FUNCTION_BLOCK Sensor_Generico_HMI (* Service Interface Function Block Type *)
  (* Standard: 61499-2 *)
  (* Version 1.6, 12/11/2026, Hidryco, Hidryco, 1.6: STS_CODIGO_ERRO, STS_CODIGO_AVISO e STS_ALM_AVISO_EST (aviso/erro do proprio dispositivo). 1.5: CommonError, Reliability e DaysToMaintenance para a IO List da Nereda. 1.4: STS_LIMITE_HH..LL (limites dos alarmes em unidade de engenharia) para o grafico. IHM do Sensor_Generico *)
  PACKAGE Hidryco.HidrycoLib;
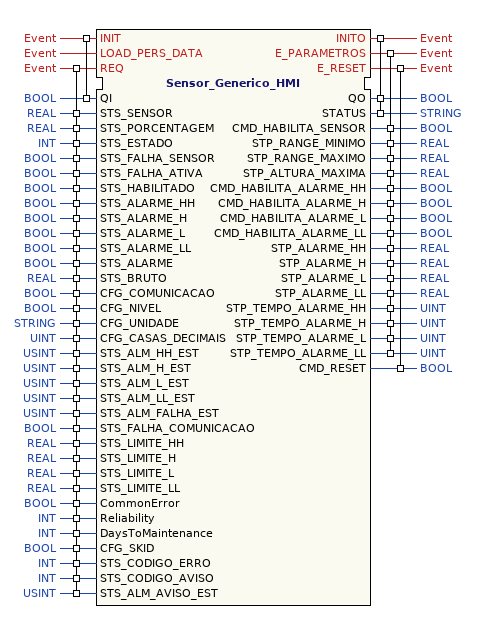
  EVENT_INPUT
    INIT WITH QI;
    LOAD_PERS_DATA; (* Reenvia os parametros persistentes *)
    REQ WITH STS_SENSOR, STS_PORCENTAGEM, STS_ESTADO, STS_FALHA_SENSOR, STS_FALHA_ATIVA, STS_HABILITADO, STS_ALARME_HH, STS_ALARME_H, STS_ALARME_L, STS_ALARME_LL, STS_ALARME, STS_BRUTO, CFG_COMUNICACAO, CFG_NIVEL, CFG_UNIDADE, CFG_CASAS_DECIMAIS, STS_ALM_HH_EST, STS_ALM_H_EST, STS_ALM_L_EST, STS_ALM_LL_EST, STS_ALM_FALHA_EST, STS_FALHA_COMUNICACAO, STS_LIMITE_HH, STS_LIMITE_H, STS_LIMITE_L, STS_LIMITE_LL, CommonError, Reliability, DaysToMaintenance, CFG_SKID, STS_CODIGO_ERRO, STS_CODIGO_AVISO, STS_ALM_AVISO_EST; (* Atualizacao de status *)
  END_EVENT
  EVENT_OUTPUT
    INITO WITH QO, STATUS;
    E_PARAMETROS WITH CMD_HABILITA_SENSOR, STP_RANGE_MINIMO, STP_RANGE_MAXIMO, STP_ALTURA_MAXIMA, CMD_HABILITA_ALARME_HH, CMD_HABILITA_ALARME_H, CMD_HABILITA_ALARME_L, CMD_HABILITA_ALARME_LL, STP_ALARME_HH, STP_ALARME_H, STP_ALARME_L, STP_ALARME_LL, STP_TEMPO_ALARME_HH, STP_TEMPO_ALARME_H, STP_TEMPO_ALARME_L, STP_TEMPO_ALARME_LL;
    E_RESET WITH CMD_RESET;
  END_EVENT
  VAR_INPUT
    QI : BOOL;
    STS_SENSOR : REAL; (* Valor em unidade de engenharia *) {SET_ATTRIBUTE(Runtime.History.Depth, 500)} {SET_ATTRIBUTE(Runtime.History.SmoothTime, 60000)} {SET_ATTRIBUTE(Runtime.History.SmoothValue, 0.1)}
    STS_PORCENTAGEM : REAL; (* Nivel em % (so sensor de nivel) *)
    STS_ESTADO : INT; (* 0 normal, 1 alerta, 2 alarme, 3 falha, 4 desabilitado *)
    STS_FALHA_SENSOR : BOOL; (* Falha do sensor (4-20 mA fora da faixa ou falha do instrumento), sem a falha de comunicacao *)
    STS_FALHA_ATIVA : BOOL; (* Qualquer falha ativa (sensor ou comunicacao) *)
    STS_HABILITADO : BOOL; (* Sensor habilitado *)
    STS_ALARME_HH : BOOL; (* Alarme HH *)
    STS_ALARME_H : BOOL; (* Alarme H *)
    STS_ALARME_L : BOOL; (* Alarme L *)
    STS_ALARME_LL : BOOL; (* Alarme LL *)
    STS_ALARME : BOOL; (* Algum alarme *)
    STS_BRUTO : REAL; (* Valor bruto lido (diagnostico) *)
    CFG_COMUNICACAO : BOOL; (* Configuracao: valor por comunicacao *)
    CFG_NIVEL : BOOL; (* Configuracao: sensor de nivel (mostra %) *)
    CFG_UNIDADE : STRING; (* Configuracao: unidade de engenharia *)
    CFG_CASAS_DECIMAIS : UINT; (* Configuracao: casas decimais *)
    STS_ALM_HH_EST : USINT; (* Estado do ALARM_BIT HH (0 normal, 1 ativo reconhecido, 2 ativo nao reconhecido, 3 saiu nao reconhecido, 4 ativo e saiu nao reconhecido) *)
    STS_ALM_H_EST : USINT; (* Estado do ALARM_BIT H (0 normal, 1 ativo reconhecido, 2 ativo nao reconhecido, 3 saiu nao reconhecido, 4 ativo e saiu nao reconhecido) *)
    STS_ALM_L_EST : USINT; (* Estado do ALARM_BIT L (0 normal, 1 ativo reconhecido, 2 ativo nao reconhecido, 3 saiu nao reconhecido, 4 ativo e saiu nao reconhecido) *)
    STS_ALM_LL_EST : USINT; (* Estado do ALARM_BIT LL (0 normal, 1 ativo reconhecido, 2 ativo nao reconhecido, 3 saiu nao reconhecido, 4 ativo e saiu nao reconhecido) *)
    STS_ALM_FALHA_EST : USINT; (* Estado do ALARM_BIT FALHA (0 normal, 1 ativo reconhecido, 2 ativo nao reconhecido, 3 saiu nao reconhecido, 4 ativo e saiu nao reconhecido) *)
    STS_FALHA_COMUNICACAO : BOOL; (* Falha de comunicacao do sensor *)
    STS_LIMITE_HH : REAL; (* Limite do alarme HH em unidade de engenharia *) {SET_ATTRIBUTE(Runtime.History.Depth, 100)} {SET_ATTRIBUTE(Runtime.History.SmoothTime, 60000)} {SET_ATTRIBUTE(Runtime.History.SmoothValue, 0)}
    STS_LIMITE_H : REAL; (* Limite do alarme H em unidade de engenharia *) {SET_ATTRIBUTE(Runtime.History.Depth, 100)} {SET_ATTRIBUTE(Runtime.History.SmoothTime, 60000)} {SET_ATTRIBUTE(Runtime.History.SmoothValue, 0)}
    STS_LIMITE_L : REAL; (* Limite do alarme L em unidade de engenharia *) {SET_ATTRIBUTE(Runtime.History.Depth, 100)} {SET_ATTRIBUTE(Runtime.History.SmoothTime, 60000)} {SET_ATTRIBUTE(Runtime.History.SmoothValue, 0)}
    STS_LIMITE_LL : REAL; (* Limite do alarme LL em unidade de engenharia *) {SET_ATTRIBUTE(Runtime.History.Depth, 100)} {SET_ATTRIBUTE(Runtime.History.SmoothTime, 60000)} {SET_ATTRIBUTE(Runtime.History.SmoothValue, 0)}
    CommonError : BOOL; (* Nereda: erro do sensor (= STS_FALHA_SENSOR) *)
    Reliability : INT; (* Nereda: confiabilidade do sensor (%), fixo em 80 *)
    DaysToMaintenance : INT; (* Nereda: dias para a manutencao (sem fonte: 0) *)
    CFG_SKID : BOOL; (* Configuracao: valor ja escalado no skid (sem ajuste de escala na IHM) *)
    STS_CODIGO_ERRO : INT; (* Codigo de erro do proprio dispositivo (0 = nenhum) *)
    STS_CODIGO_AVISO : INT; (* Codigo de aviso do proprio dispositivo (0 = nenhum) *)
    STS_ALM_AVISO_EST : USINT; (* Estado do ALARM_BIT de aviso do dispositivo (0 normal, 1 ativo reconhecido, 2 ativo nao reconhecido, 3 saiu nao reconhecido, 4 ativo e saiu) *)
  END_VAR
  VAR_OUTPUT
    QO : BOOL; (* Event Output Qualifier *)
    STATUS : STRING; (* Service Status *)
    CMD_HABILITA_SENSOR : BOOL; (* Sensor habilitado *)
    STP_RANGE_MINIMO : REAL; (* Valor de engenharia em 4 mA *)
    STP_RANGE_MAXIMO : REAL; (* Valor de engenharia em 20 mA *)
    STP_ALTURA_MAXIMA : REAL; (* Altura maxima do tanque (nivel) *)
    CMD_HABILITA_ALARME_HH : BOOL; (* Alarme HH habilitado *)
    CMD_HABILITA_ALARME_H : BOOL; (* Alarme H habilitado *)
    CMD_HABILITA_ALARME_L : BOOL; (* Alarme L habilitado *)
    CMD_HABILITA_ALARME_LL : BOOL; (* Alarme LL habilitado *)
    STP_ALARME_HH : REAL; (* Setpoint do alarme HH *)
    STP_ALARME_H : REAL; (* Setpoint do alarme H *)
    STP_ALARME_L : REAL; (* Setpoint do alarme L *)
    STP_ALARME_LL : REAL; (* Setpoint do alarme LL *)
    STP_TEMPO_ALARME_HH : UINT; (* Tempo do alarme HH (s); padrao 5 s (retardo contra alarme falso, ISA-18.2) *)
    STP_TEMPO_ALARME_H : UINT; (* Tempo do alarme H (s); padrao 5 s (retardo contra alarme falso, ISA-18.2) *)
    STP_TEMPO_ALARME_L : UINT; (* Tempo do alarme L (s); padrao 5 s (retardo contra alarme falso, ISA-18.2) *)
    STP_TEMPO_ALARME_LL : UINT; (* Tempo do alarme LL (s); padrao 5 s (retardo contra alarme falso, ISA-18.2) *)
    CMD_RESET : BOOL; (* Reset de falha e alarmes *)
  END_VAR
  SERVICE /
    SEQUENCE 
    END_SEQUENCE
  END_SERVICE
END_FUNCTION_BLOCK
